FUNCTION_BLOCK LowestRecipeElapsedTime (* Basic Function Block Type *)
  (* Standard: 61499-2 *)
  (* Version 0.0, 10/6/2026, Schneider Electric, Template *)
  PACKAGE SE.Nereda;
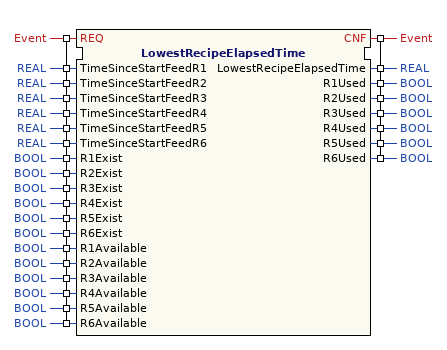
  EVENT_INPUT
    REQ WITH TimeSinceStartFeedR1, TimeSinceStartFeedR2, TimeSinceStartFeedR3, TimeSinceStartFeedR4, TimeSinceStartFeedR5, TimeSinceStartFeedR6, R1Exist, R2Exist, R3Exist, R4Exist, R5Exist, R6Exist, R1Available, R2Available, R3Available, R4Available, R5Available, R6Available; (* Normal Execution Request *)
  END_EVENT
  EVENT_OUTPUT
    CNF WITH LowestRecipeElapsedTime, R1Used, R2Used, R3Used, R4Used, R5Used, R6Used; (* Execution Confirmation *)
  END_EVENT
  VAR_INPUT
    TimeSinceStartFeedR1 : REAL;
    TimeSinceStartFeedR2 : REAL;
    TimeSinceStartFeedR3 : REAL;
    TimeSinceStartFeedR4 : REAL;
    TimeSinceStartFeedR5 : REAL;
    TimeSinceStartFeedR6 : REAL;
    R1Exist : BOOL;
    R2Exist : BOOL;
    R3Exist : BOOL;
    R4Exist : BOOL;
    R5Exist : BOOL;
    R6Exist : BOOL;
    R1Available : BOOL;
    R2Available : BOOL;
    R3Available : BOOL;
    R4Available : BOOL;
    R5Available : BOOL;
    R6Available : BOOL;
  END_VAR
  VAR_OUTPUT
    LowestRecipeElapsedTime : REAL;
    R1Used : BOOL;
    R2Used : BOOL;
    R3Used : BOOL;
    R4Used : BOOL;
    R5Used : BOOL;
    R6Used : BOOL;
  END_VAR
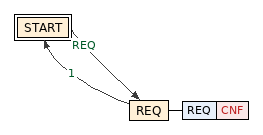
  EC_STATES
    START; (* Initial State *)
    REQ : REQ -> CNF; (* Normal execution *)
  END_STATES
  EC_TRANSITIONS
    START TO REQ := REQ;
    REQ TO START := 1;
  END_TRANSITIONS
  ALGORITHM REQ IN ST: (* Normally executed algorithm *)
;
//R1Used := R1Exist AND R1Available;
//R2Used := R2Exist AND R2Available;
//R3Used := R3Exist AND R3Available;
//R4Used := R4Exist AND R4Available;
//R5Used := R5Exist AND R5Available;
//R6Used := R6Exist AND R6Available;

R1Used := R1Exist;
R2Used := R2Exist;
R3Used := R3Exist;
R4Used := R4Exist;
R5Used := R5Exist;
R6Used := R6Exist;


// Initialize with the first used reactor
IF R1Used THEN
    LowestRecipeElapsedTime := TimeSinceStartFeedR1;

ELSIF R2Used THEN
    LowestRecipeElapsedTime := TimeSinceStartFeedR2;

ELSIF R3Used THEN
    LowestRecipeElapsedTime := TimeSinceStartFeedR3;

ELSIF R4Used THEN
    LowestRecipeElapsedTime := TimeSinceStartFeedR4;

ELSIF R5Used THEN
    LowestRecipeElapsedTime := TimeSinceStartFeedR5;

ELSIF R6Used THEN
    LowestRecipeElapsedTime := TimeSinceStartFeedR6;

END_IF;


// Find the lowest value
IF R1Used AND (TimeSinceStartFeedR1 < LowestRecipeElapsedTime) THEN
    LowestRecipeElapsedTime := TimeSinceStartFeedR1;
END_IF;

IF R2Used AND (TimeSinceStartFeedR2 < LowestRecipeElapsedTime) THEN
    LowestRecipeElapsedTime := TimeSinceStartFeedR2;
END_IF;

IF R3Used AND (TimeSinceStartFeedR3 < LowestRecipeElapsedTime) THEN
    LowestRecipeElapsedTime := TimeSinceStartFeedR3;
END_IF;

IF R4Used AND (TimeSinceStartFeedR4 < LowestRecipeElapsedTime) THEN
    LowestRecipeElapsedTime := TimeSinceStartFeedR4;
END_IF;

IF R5Used AND (TimeSinceStartFeedR5 < LowestRecipeElapsedTime) THEN
    LowestRecipeElapsedTime := TimeSinceStartFeedR5;
END_IF;

IF R6Used AND (TimeSinceStartFeedR6 < LowestRecipeElapsedTime) THEN
    LowestRecipeElapsedTime := TimeSinceStartFeedR6;
END_IF;
  END_ALGORITHM
END_FUNCTION_BLOCK
